{attribute 'qualified_only'}
{attribute 'strict'}
{attribute 'to_string'}
TYPE E_LEDs :
(
	NONE := 0,
    START_BTN := 1,
    STOP_BTN := 2,
    RESET_BTN := 3
);
END_TYPE

(* stored: Version 1.1.0.1
   DUT E_LEDs: Id {fc31990f-c939-4669-9b6b-fb72d46ae7d7} *)
